Staubli VAL3: main.pgx

program main()
begin
  close(tCurrentTool)
  pPointRs.config.shoulder = lefty
  pPointRs2.config.shoulder = lefty
  mCurrentSpeed.tvel = 100.00
  mCurrentSpeed.blend = joint
  mCurrentSpeed.reach = 0.010
  mCurrentSpeed.leave = 0.010
  // Program EdgeProg start
  // Program generated by RoboDK v6.0.7 for Staubli TS20 FL 100 TC on XX/XX/XXXX 18:00:00
  // Using nominal kinematics.
  mCurrentSpeed.tvel = 123.456
  mCurrentSpeed.reach = -1.000
  mCurrentSpeed.leave = -1.000
  call MoveJoint(-15.00000,40.00000,20.00000,90.00000)
  mCurrentSpeed.reach = 12.500
  mCurrentSpeed.leave = 12.500
  call MoveLine(-624.230,571.208,454.620,81.604,51.756,-128.588)
  delay(0.000)
  delay(1.234)
  popUpMsg("A long message with "quotes", 'apostrophes' & symbols: <>[]{}()=+-*/%;#@! and more text to make it longer than eighty characters")
  // Comment with ; semicolon
  Gripper=ON
  Output[12]=false
  Pressure=true
  watch(PartPresent==true,250.0)
  watch(Input[7]==1)
  //call prog:Do Something(1, 2)
  x = 1
  call MoveJoint(30.00000,25.00000,80.00000,-45.00000)

  waitEndMove()
  // Program EdgeProg end

end
